(* PLC project Motor_StartStop_TM241CE24T, PLCAutoPilot M241 Generator 2.0 *)
(* stored: creationDateTime 2025-12-30T00:00:00, modificationDateTime 2025-12-30T00:00:00 *)

(* Motor Start/Stop Control Program Features: - 3 second startup delay (anti-chatter) - Overload fault latching with automatic reset - Emergency stop interlock - Run and fault indication lamps Safety: - StopPB is NC (fail-safe: wire break = motor stops) - EmergencyStop is NC (fail-safe) - OverloadTrip is NC (fail-safe) Generated by PLCAutoPilot for TM241CE24T *)
PROGRAM Motor_Control
  VAR
    StartPB : BOOL;  (* Start Pushbutton (NO) - %IX0.0 *)
    StopPB : BOOL;  (* Stop Pushbutton (NC) - %IX0.1 *)
    OverloadTrip : BOOL;  (* Thermal Overload (NC) - %IX0.2 *)
    EmergencyStop : BOOL;  (* E-Stop (NC) - %IX0.3 *)
    MotorContactor : BOOL;  (* Main Contactor - %QX0.0 *)
    RunIndicator : BOOL;  (* Run Lamp - %QX0.1 *)
    FaultIndicator : BOOL;  (* Fault Lamp - %QX0.2 *)
    MotorRunning : BOOL;
    MotorFault : BOOL;
    SafetyOK : BOOL;
    StartupTimer : TON;
  END_VAR

            
// ============================================
// MOTOR START/STOP CONTROL
// TM241CE24T - PLCAutoPilot Generated
// ============================================
//
// I/O MAPPING:
// Inputs:
//   StartPB       - %IX0.0 (NO pushbutton)
//   StopPB        - %IX0.1 (NC pushbutton)
//   OverloadTrip  - %IX0.2 (NC thermal relay)
//   EmergencyStop - %IX0.3 (NC E-Stop)
//
// Outputs:
//   MotorContactor - %QX0.0 (Main contactor K1)
//   RunIndicator   - %QX0.1 (Run lamp)
//   FaultIndicator - %QX0.2 (Fault lamp)
// ============================================

// Read physical inputs (assign I/O addresses in GVL)
// StartPB := %IX0.0;
// StopPB := %IX0.1;
// OverloadTrip := %IX0.2;
// EmergencyStop := %IX0.3;

// Safety interlock check
// E-Stop must be OK (NC contact = TRUE when OK)
// Overload must be OK (NC contact = TRUE when OK)
SafetyOK := EmergencyStop AND NOT OverloadTrip;

// Fault latching
// Set fault when overload trips
// Reset fault when Start is pressed AND overload is cleared
IF OverloadTrip THEN
    MotorFault := TRUE;
END_IF;

IF StartPB AND NOT OverloadTrip THEN
    MotorFault := FALSE;
END_IF;

// Startup timer (3 second anti-chatter delay)
// Timer runs when Start pressed, Safety OK, and no fault
StartupTimer(
    IN := StartPB AND SafetyOK AND NOT MotorFault AND NOT MotorRunning,
    PT := T#3S
);

// Motor running logic
// SET: Timer complete (3 seconds of continuous Start press)
IF StartupTimer.Q THEN
    MotorRunning := TRUE;
END_IF;

// RESET: Stop pressed OR Safety NOT OK OR Fault
IF NOT StopPB OR NOT SafetyOK OR MotorFault THEN
    MotorRunning := FALSE;
END_IF;

// Write to outputs
MotorContactor := MotorRunning;
RunIndicator := MotorRunning;
FaultIndicator := MotorFault;

// Write to physical outputs (assign I/O addresses in GVL)
// %QX0.0 := MotorContactor;
// %QX0.1 := RunIndicator;
// %QX0.2 := FaultIndicator;
            
          
END_PROGRAM

CONFIGURATION TM241CE24T
  RESOURCE Application ON PLC
    TASK MAST(INTERVAL := T#20ms, PRIORITY := 1);
    PROGRAM Motor_Control_Inst WITH MAST : Motor_Control;
  END_RESOURCE
END_CONFIGURATION
